Universal Robots URScript: T007_qwen2.5-coder_32b-instruct-q4_0_baseline_rep1.urscript

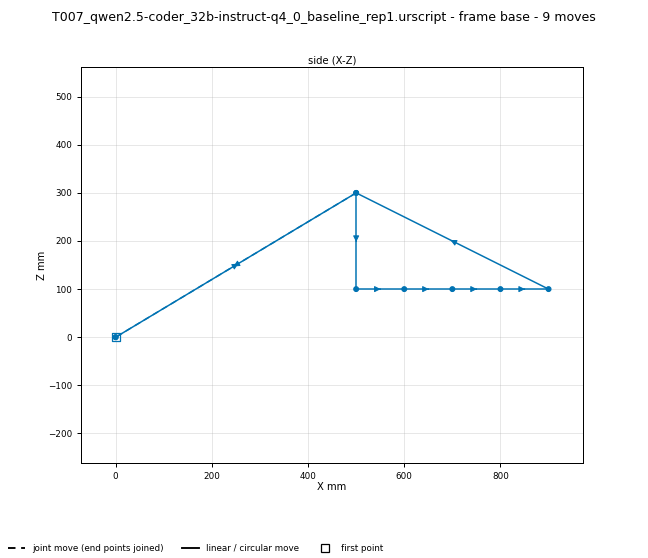
[picture p0: tool path of T007_qwen2.5-coder_32b-instruct-q4_0_baseline_rep1.urscript in frame base, 9 of 9 moves have a stored position in this frame; points joined in program order, loops and branches not executed]
# URScript for Curved Contour Weld - Hybrid Mode (T007)

# Home position
movej(p[0.0, -1.5708, 0.0, -1.5708, 0.0, 0.0], a=1.2, v=1.2)

# Approach above weld fixture
movel(p[0.5, -1.5708, 0.3, -1.5708, 0.0, 0.0], a=1.2, v=1.0)

# Descend to weld start
movel(p[0.5, -1.5708, 0.1, -1.5708, 0.0, 0.0], a=1.2, v=0.4)

# Weld midpoint
movel(p[0.6, -1.5708, 0.1, -1.5708, 0.0, 0.0], a=1.2, v=0.2)

# Weld end
movel(p[0.7, -1.5708, 0.1, -1.5708, 0.0, 0.0], a=1.2, v=0.2)

# Continue weld path (2 more points)
movel(p[0.8, -1.5708, 0.1, -1.5708, 0.0, 0.0], a=1.2, v=0.2)
movel(p[0.9, -1.5708, 0.1, -1.5708, 0.0, 0.0], a=1.2, v=0.2)

# Return to approach position
movel(p[0.5, -1.5708, 0.3, -1.5708, 0.0, 0.0], a=1.2, v=1.0)

# Return to home position
movej(p[0.0, -1.5708, 0.0, -1.5708, 0.0, 0.0], a=1.2, v=1.2)
